Fanuc KAREL source: KT00599.KL

PROGRAM KT00599
%NOLOCKGROUP
VAR
  I1: INTEGER
  I2: INTEGER
  OUT: REAL
BEGIN
  I1 = 2
  I2 = 3
  I1 = 2
  I2 = 3
  OUT = NOT I1
END KT00599
